// Argument container. Values are stored as text, ready for the formatter.
FUNCTION_BLOCK FB_EventArgs IMPLEMENTS I_ArgumentBuilder, I_ArgumentSource
VAR
	aValues	: ARRAY[0..GVL_EventFramework.cMaxArguments - 1] OF T_MaxString;
	nCount	: USINT;
END_VAR

METHOD PRIVATE Append : I_ArgumentBuilder
VAR_INPUT
	sValue	: T_MaxString;
END_VAR
IF nCount < GVL_EventFramework.cMaxArguments THEN
	aValues[nCount] := sValue;
	nCount := nCount + 1;
END_IF
Append := THIS^;
END_METHOD

METHOD Clear : I_ArgumentBuilder
nCount := 0;
Clear := THIS^;
END_METHOD

METHOD AddString : I_ArgumentBuilder
VAR_INPUT
	sValue	: T_MaxString;
END_VAR
AddString := Append(sValue);
END_METHOD

METHOD AddDInt : I_ArgumentBuilder
VAR_INPUT
	nValue	: DINT;
END_VAR
AddDInt := Append(DINT_TO_STRING(nValue));
END_METHOD

METHOD AddLReal : I_ArgumentBuilder
VAR_INPUT
	fValue		: LREAL;
	nDecimals	: USINT;	// 0..9
END_VAR
VAR
	nDigits	: USINT;
	nScale	: LINT := 1;
	nScaled	: LINT;
	i		: USINT;
	sFrac	: STRING(20);
	sValue	: T_MaxString;
END_VAR
nDigits := MIN(nDecimals, 9);
FOR i := 1 TO nDigits DO
	nScale := nScale * 10;
END_FOR

// Fixed-point formatting avoids LREAL_TO_STRING artefacts like 82.350000000000009
nScaled := LREAL_TO_LINT(ABS(fValue) * LINT_TO_LREAL(nScale));
sValue := LINT_TO_STRING(nScaled / nScale);
IF nDigits > 0 THEN
	sFrac := LINT_TO_STRING(nScaled MOD nScale);
	WHILE LEN(sFrac) < nDigits DO
		sFrac := CONCAT('0', sFrac);
	END_WHILE
	sValue := CONCAT(CONCAT(sValue, '.'), sFrac);
END_IF
IF fValue < 0 AND nScaled <> 0 THEN
	sValue := CONCAT('-', sValue);
END_IF

AddLReal := Append(sValue);
END_METHOD

METHOD AddBool : I_ArgumentBuilder
VAR_INPUT
	bValue	: BOOL;
END_VAR
IF bValue THEN
	AddBool := Append('TRUE');
ELSE
	AddBool := Append('FALSE');
END_IF
END_METHOD

METHOD GetArgument : T_MaxString
VAR_INPUT
	nIndex	: USINT;
END_VAR
IF nIndex < nCount THEN
	GetArgument := aValues[nIndex];
END_IF
END_METHOD

PROPERTY Count : USINT
GET
Count := nCount;
END_GET
END_PROPERTY

END_FUNCTION_BLOCK

(* stored: Version 1.1.0.1, ProductVersion 3.1.4026.26
   POU FB_EventArgs: Id {9557b18b-aeea-4a94-882b-d4ef219de25c}, SpecialFunc None
   Method Append: Id {5822f03d-3d66-4104-8b26-0bce187fbd25}
   Method Clear: Id {fa4bebbe-5a70-49b5-ae94-66d822ae4a95}
   Method AddString: Id {6321ec74-47a3-4560-8567-62c49383d67a}
   Method AddDInt: Id {aab139e2-707b-432c-82bb-de1b60a37026}
   Method AddLReal: Id {eb8b8006-a215-4b79-bc9b-c1a52446d4b6}
   Method AddBool: Id {50546d3a-aa62-4e4a-804b-496d49daa64c}
   Method GetArgument: Id {e47617db-6390-44ce-92d7-49cfe754980a}
   Property Count: Id {5e716aa1-3895-4f9a-b599-bb2637a2593e}
   Get Get: Id {0e5c7045-84fd-4ab3-8181-21fc4f575266} *)
